(* IEC 61131-3 sources: SortJet_MasterSPS_Aufbau.fbsproj/08_POUs/Basis Programmbausteine/StartUpCheck.prg.st^, 11 files *)

(* ---- checkAchsID.meth.st ---- *)
(* METADATA
{
	"v3Meta": {
		"objectGuid": "61da6f1d-6d44-4478-83af-d8c1dc57ab14"
	}
}
*)
METHOD checkAchsID
VAR_INPUT
  wAchsID : REFERENCE TO WORD;
END_VAR
VAR
  cLOG_HANDLE : RTS_IEC_HANDLE := RTS_INVALID_HANDLE;
END_VAR
IF NOT __ISVALIDREF(wAchsID) THEN
  RETURN;
END_IF

IF wAchsID = 65 THEN
  RETURN; // explizit erlaubt
END_IF;

IF wAchsID > 65 THEN
  CmpLog.LogAdd2(cLOG_HANDLE, 16#00010000, 16#00000001, 16#00000010, 0, 'Konfigurationsfehler: Konfigurierte AchsID zu groß');
  SysExceptGenerateException(RtsExceptions.RTSEXCPT_NONCONTINUABLE); // AchsID ist zu groß
  NullRef := TRUE; // Falls die obenstehende Exception nicht auslöst, auf eine NullReferenz zugreifen -> Exception auch in Simulation.
END_IF

IF aUsedAchsIDs[wAchsID] THEN
  CmpLog.LogAdd2(cLOG_HANDLE, 16#00010000, 16#00000001, 16#00000010, 0, 'Konfigurationsfehler: AchsID mehrfach vergeben');
  SysExceptGenerateException(RtsExceptions.RTSEXCPT_NONCONTINUABLE); // AchsID bereits in benutzung!
  NullRef := TRUE; // Falls die obenstehende Exception nicht auslöst, auf eine NullReferenz zugreifen -> Exception auch in Simulation.
END_IF

aUsedAchsIDs[wAchsID] := TRUE;
END_METHOD

(* ---- checkAutomatikkreis.meth.st ---- *)
(* METADATA
{
	"v3Meta": {
		"objectGuid": "b3622f19-1aaf-4182-891a-040c2736cdb4"
	}
}
*)
METHOD checkAutomatikkreis
VAR_INPUT
  Basis : REFERENCE TO StationBasisParameter_ST;
END_VAR
VAR
  x : WORD;
  bAutomatikkreisGefunden : BOOL;
  eaAutomatikkreis : ARRAY [cERSTER_AUTOMATIKKREIS..cANZAHL_AUTOMATIKKREISE] OF BOOL;
END_VAR

// eaAutomatikkreis prüfen - mindestens ein AK muss gesetzt sein und nur vorhandene Automatikkreise dürfen gesetzt sein

bAutomatikkreisGefunden := FALSE;

FOR x := cERSTER_AUTOMATIKKREIS TO cANZAHL_AUTOMATIKKREISE DO
  IF Basis.stMKs.eaAutomatikkreis[x] <> 0 THEN
    bAutomatikkreisGefunden := TRUE;
  END_IF
END_FOR
IF NOT bAutomatikkreisGefunden THEN
  CmpLog.LogAdd2(cLOG_HANDLE, 16#00010000, 16#00000001, 16#00000010, 0, 'Kein Automatikkreis konfiguriert');
  SysExceptGenerateException(RtsExceptions.RTSEXCPT_NONCONTINUABLE);
  NullRef := TRUE;
END_IF

FOR x := cERSTER_AUTOMATIKKREIS TO cANZAHL_AUTOMATIKKREISE DO
  IF Basis.stMKs.eaAutomatikkreis[x] <> 0 THEN
    IF ( Basis.stMKs.eaAutomatikkreis[x] < cERSTER_AUTOMATIKKREIS ) OR ( Basis.stMKs.eaAutomatikkreis[x] > cLETZTER_AUTOMATIKKREIS ) THEN
      CmpLog.LogAdd2(cLOG_HANDLE, 16#00010000, 16#00000001, 16#00000010, Basis.stMKs.eaAutomatikkreis[x], 'Automatikkreis existiert nicht');
      SysExceptGenerateException(RtsExceptions.RTSEXCPT_NONCONTINUABLE);
      NullRef := TRUE;
    END_IF
  END_IF
END_FOR
END_METHOD

(* ---- checkAutomatikkreiseMK.meth.st ---- *)
(* METADATA
{
	"v3Meta": {
		"objectGuid": "4f81610e-119d-462b-b6ef-1c5c06c97f10"
	}
}
*)
METHOD checkAutomatikkreiseMK
VAR_INPUT
END_VAR
VAR
  x : WORD;
END_VAR
FOR x := cERSTER_AUTOMATIKKREIS TO cLETZTER_AUTOMATIKKREIS DO
  IF apgMKAutomatikkreise[x].epAutomatikkreis_Transfershuttle = 0 THEN
    CmpLog.LogAdd2(cLOG_HANDLE, 16#00010000, 16#00000001, 16#00000040, x, 'apgMKAutomatikkreise: Automatikkreis nicht definiert');
    SysExceptGenerateException(RtsExceptions.RTSEXCPT_NONCONTINUABLE);
    NullRef := TRUE;
  END_IF
END_FOR
END_METHOD

(* ---- checkDurchgaenge.meth.st ---- *)
(* METADATA
{
	"v3Meta": {
		"objectGuid": "22b8b65b-6376-41dd-ab5a-bf0c9c2eeadd"
	}
}
*)
METHOD checkDurchgaenge
VAR_INPUT
END_VAR
VAR
  x : WORD;
END_VAR

FOR x := cERSTER_DURCHGANG TO cANZAHL_DURCHGANGE DO
  IF apgMKDurchgang[x].eDurchgang = 0 THEN
    CmpLog.LogAdd2(cLOG_HANDLE, 16#00010000, 16#00000001, 16#00000060, x, 'apgMKDurchgang: Durchgang nicht definiert');
    SysExceptGenerateException(RtsExceptions.RTSEXCPT_NONCONTINUABLE);
    NullRef := TRUE;
  END_IF
END_FOR
END_METHOD

(* ---- checkGlastransportOptionen.meth.st ---- *)
(* METADATA
{
	"v3Meta": {
		"objectGuid": "9d81c253-8159-4cb9-9043-a22c56ba0597"
	}
}
*)
METHOD checkGlastransportOptionen
VAR_INPUT
  Basis                : REFERENCE TO StationBasisParameter_ST;
  bAustransportPruefen : BOOL; // Austransport-Option wird nur vom Shuttle (Vorab) gebraucht
END_VAR
VAR
  n : WORD;
END_VAR

// Lage der letzten Scheibe im Eintransport (eGlastransport) muss je konfiguriertem Partner gesetzt sein,
// im Austransport nur beim Shuttle (Vorab). Transfershuttle als Partner hat die Option nicht.
// eGlastransport_Default gilt als fehlende Konfiguration, die SPS bleibt stehen.
FOR n := cERSTES_SHUTTLE TO cLETZTE_FREMDANLAGE_EINLAUF DO

  IF (     ( Basis.stMKs.stSchnittstellendaten.aEintransporte.Station[n] <> TransportRichtung_EN.Default )
       AND NOT ( ( n >= cERSTES_TRANSFERSHUTTLE ) AND ( n <= cLETZTES_TRANSFERSHUTTLE ) )
       AND ( Basis.stMKs.stSchnittstellendaten.aEintransporte.Glastransport[n] = eGlastransport_Default ) )
  THEN
    CmpLog.LogAdd2(cLOG_HANDLE, 16#00010000, 16#00000001, 16#00000010, 0, 'aEintransporte.Glastransport darf bei konfiguriertem Partner nicht Default sein');
    SysExceptGenerateException(RtsExceptions.RTSEXCPT_NONCONTINUABLE);
    NullRef := TRUE;
  END_IF

  IF (     bAustransportPruefen
       AND ( Basis.stMKs.stSchnittstellendaten.aAustransporte.Station[n] <> TransportRichtung_EN.Default )
       AND ( Basis.stMKs.stSchnittstellendaten.aAustransporte.Glastransport[n] = eGlastransport_Default ) )
  THEN
    CmpLog.LogAdd2(cLOG_HANDLE, 16#00010000, 16#00000001, 16#00000010, 0, 'aAustransporte.Glastransport darf bei konfiguriertem Partner nicht Default sein');
    SysExceptGenerateException(RtsExceptions.RTSEXCPT_NONCONTINUABLE);
    NullRef := TRUE;
  END_IF

END_FOR
END_METHOD

(* ---- checkMeldungsnummer.meth.st ---- *)
(* METADATA
{
	"v3Meta": {
		"objectGuid": "b642c49f-6ffa-4fce-b10f-dd7fb5dad387"
	}
}
*)
METHOD checkMeldungsnummer
VAR_INPUT
  Basis : REFERENCE TO StationBasisParameter_ST;
END_VAR

// wMeldungsnummer prüfen - nicht 0 und nicht doppelt vergeben
IF Basis.stMKs.wMeldungsnummer = 0 THEN
  CmpLog.LogAdd2(cLOG_HANDLE, 16#00010000, 16#00000001, 16#00000010, 0, 'wMeldungsnummer darf nicht 0 sein');
  SysExceptGenerateException(RtsExceptions.RTSEXCPT_NONCONTINUABLE);
  NullRef := TRUE;
END_IF
IF aUsedMeldungsnummern[Basis.stMKs.wMeldungsnummer] THEN
  CmpLog.LogAdd2(cLOG_HANDLE, 16#00010000, 16#00000001, 16#00000010, 0, 'wMeldungsnummer mehrfach konfiguriert');
  SysExceptGenerateException(RtsExceptions.RTSEXCPT_NONCONTINUABLE);
  NulLRef := TRUE;
END_IF
aUsedMeldungsnummern[Basis.stMKs.wMeldungsnummer] := TRUE;
END_METHOD

(* ---- checkMKVerfahrparameter.meth.st ---- *)
(* METADATA
{
	"v3Meta": {
		"objectGuid": "c7964ec2-357c-46cb-95df-ee4bc270f3f8"
	}
}
*)
METHOD checkMKVerfahrparameter
VAR_INPUT
END_VAR
VAR
  x : WORD;
END_VAR

FOR x := cERSTES_SHUTTLE TO cLETZTES_SHUTTLE DO
  IF ( apgShuttleVerfahrparameter[x].eParkposition = 0 ) THEN
    CmpLog.LogAdd2(cLOG_HANDLE, 16#00010000, 16#00000001, 16#00000020, 0, 'apgShuttleVerfahrparameter steht auf Default');
    SysExceptGenerateException(RtsExceptions.RTSEXCPT_NONCONTINUABLE);
    NullRef := TRUE;
  END_IF
END_FOR
FOR x := cERSTES_TRANSFERSHUTTLE TO cLETZTES_TRANSFERSHUTTLE DO
  IF ( apgTransfershuttleVerfahrparameter[x].eParkposition = 0 ) THEN
    CmpLog.LogAdd2(cLOG_HANDLE, 16#00010000, 16#00000001, 16#00000021, 0, 'apgTransfershuttleVerfahrparameter steht auf Default');
    SysExceptGenerateException(RtsExceptions.RTSEXCPT_NONCONTINUABLE);
    NullRef := TRUE;
  END_IF
END_FOR
END_METHOD

(* ---- checkSicherheitskreiseMK.meth.st ---- *)
(* METADATA
{
	"v3Meta": {
		"objectGuid": "1e7d8eb1-23f2-478f-a0da-97a7b6d734ce"
	}
}
*)
METHOD checkSicherheitskreiseMK
VAR_INPUT
END_VAR
VAR
  x : WORD;
END_VAR

FOR x := cERSTER_SICHERHEITSKREIS TO cLETZTER_SICHERHEITSKREIS DO
  IF apgMKSicherheiskreis[x].eSicherheitskreis = 0 THEN
    CmpLog.LogAdd2(cLOG_HANDLE, 16#00010000, 16#00000001, 16#00000050, x, 'apgMKSicherheiskreis: Sicherheitskreis nicht definiert');
    SysExceptGenerateException(RtsExceptions.RTSEXCPT_NONCONTINUABLE);
    NullRef := TRUE;
  END_IF
END_FOR
END_METHOD

(* ---- checkStationsnummern.meth.st ---- *)
(* METADATA
{
	"v3Meta": {
		"objectGuid": "577e9539-3133-4f06-80f9-5ab9a23fcb59"
	}
}
*)
METHOD checkStationsnummern
VAR_INPUT
  Basis : REFERENCE TO StationBasisParameter_ST;
END_VAR

// stStationsNummern prüfen - keine 0 keine doppelt vergeben
IF Basis.stMKs.stStationsNummern.NummerIntern = 0 THEN
  CmpLog.LogAdd2(cLOG_HANDLE, 16#00010000, 16#00000001, 16#00000010, 0, 'StationsNummer Intern darf nicht 0 sein');
  SysExceptGenerateException(RtsExceptions.RTSEXCPT_NONCONTINUABLE);
  NullRef := TRUE;
END_IF
IF aUsedStationNrIntern[Basis.stMKs.stStationsNummern.NummerIntern] THEN
  CmpLog.LogAdd2(cLOG_HANDLE, 16#00010000, 16#00000001, 16#00000010, 0, 'StationsNummer Intern doppelt vergeben');
  SysExceptGenerateException(RtsExceptions.RTSEXCPT_NONCONTINUABLE);
  NullRef := TRUE;
END_IF
aUsedStationNrIntern[Basis.stMKs.stStationsNummern.NummerIntern] := TRUE;

IF Basis.stMKs.stStationsNummern.NummerSPS = 0 THEN
  CmpLog.LogAdd2(cLOG_HANDLE, 16#00010000, 16#00000001, 16#00000010, 0, 'StationsNummer SPS darf nicht 0 sein');
  SysExceptGenerateException(RtsExceptions.RTSEXCPT_NONCONTINUABLE);
  NullRef := TRUE;
END_IF
IF aUsedStationNrSPS[Basis.stMKs.stStationsNummern.NummerSPS] THEN
  CmpLog.LogAdd2(cLOG_HANDLE, 16#00010000, 16#00000001, 16#00000010, 0, 'StationsNummer SPS doppelt vergeben');
  SysExceptGenerateException(RtsExceptions.RTSEXCPT_NONCONTINUABLE);
  NullRef := TRUE;
END_IF
aUsedStationNrSPS[Basis.stMKs.stStationsNummern.NummerSPS] := TRUE;

// INFO: Extern kann nicht geprüft werden, da undefinierter Nummernkreis!
END_METHOD

(* ---- checkStationsTyp.meth.st ---- *)
(* METADATA
{
	"v3Meta": {
		"objectGuid": "1787c9d8-e07d-471d-967c-af403122e309"
	}
}
*)
METHOD checkStationsTyp
VAR_INPUT
  Basis : REFERENCE TO StationBasisParameter_ST;
END_VAR

// eStationsTyp prüfen - nicht 0
IF Basis.stMKs.eStationsTyp = 0 THEN
  CmpLog.LogAdd2(cLOG_HANDLE, 16#00010000, 16#00000001, 16#00000010, 0, 'eStationsTyp darf nicht 0 sein');
  SysExceptGenerateException(RtsExceptions.RTSEXCPT_NONCONTINUABLE);
  NullRef := TRUE;
END_IF
END_METHOD

(* ---- checkZentralschmierung.meth.st ---- *)
(* METADATA
{
	"v3Meta": {
		"objectGuid": "5eb94ffc-f2d1-4fcc-9867-11fb69ff17a0"
	}
}
*)
METHOD checkZentralschmierung
VAR_INPUT
END_VAR
VAR
  x, y : WORD;
END_VAR

FOR x := cERSTES_SHUTTLE TO cLETZTES_SHUTTLE DO
  FOR y := 1 TO 2 DO
    IF apgMKShuttleZentralschmierung[x].aiAnzahlHuebe[y] = 0 THEN
      CmpLog.LogAdd2(cLOG_HANDLE, 16#00010000, 16#00000001, 16#00000030, i, 'Shuttle-Zentralschmierung: Anzahl Huebe = 0');
      SysExceptGenerateException(RtsExceptions.RTSEXCPT_NONCONTINUABLE);
      NullRef := TRUE;
    END_IF;

    IF apgMKShuttleZentralschmierung[x].adiZuFahrenderWegBisSchmierung[y] = 0 THEN
      CmpLog.LogAdd2(cLOG_HANDLE, 16#00010000, 16#00000001, 16#00000031, i, 'Shuttle-Zentralschmierung: Weg bis Schmierung = 0');
      SysExceptGenerateException(RtsExceptions.RTSEXCPT_NONCONTINUABLE);
      NullRef := TRUE;
    END_IF
  END_FOR
END_FOR

FOR x := cERSTES_TRANSFERSHUTTLE TO cLETZTES_TRANSFERSHUTTLE DO
  FOR y := 1 TO 2 DO
    IF apgMKTransfershuttleZentralschmierung[x].aiAnzahlHuebe[y] = 0 THEN
      CmpLog.LogAdd2(cLOG_HANDLE, 16#00010000, 16#00000001, 16#00000032, i, 'Transfershuttle-Zentralschmierung: Anzahl Huebe = 0');
      SysExceptGenerateException(RtsExceptions.RTSEXCPT_NONCONTINUABLE);
      NullRef := TRUE;
    END_IF;

    IF apgMKTransfershuttleZentralschmierung[x].adiZuFahrenderWegBisSchmierung[y] = 0 THEN
      CmpLog.LogAdd2(cLOG_HANDLE, 16#00010000, 16#00000001, 16#00000033, i, 'Transfershuttle-Zentralschmierung: Weg bis Schmierung = 0');
      SysExceptGenerateException(RtsExceptions.RTSEXCPT_NONCONTINUABLE);
      NullRef := TRUE;
    END_IF
  END_FOR
END_FOR
END_METHOD
